(*
SPDX-FileCopyrightText: © 2026 Oleksandr Tiutyk <trofimich@gmail.com>
SPDX-License-Identifier: MIT
License: https://opensource.org/license/mit
*)

(*!
<summary>Creates application-specific activities and conditions for Workflows.CreateElement.</summary>
<description>Invoked in the owning task during configuration. The common creation path registers a successful result.</description>
*)
INTERFACE IWorkflowElementFactory

(*!
<summary>Creates an unregistered element for a recognized qualified PLC type.</summary>
<description>Return zero for an unknown type. For a recognized type return one fresh, unattached dynamic element
associated with workflow. Transfer exclusive ownership on return. On failure clean up before propagating;
a failed allocation must raise terminal OOM. Do not register or publish the element in this callback.</description>
<param name="typeName">Case-sensitive namespace and PLC type name.</param>
<param name="workflow">Prospective owner supplied to the node constructor.</param>
*)
METHOD CreateElement : IWorkflowElement
VAR_INPUT
	typeName : STRING(255);
	workflow : IWorkflow;
END_VAR
END_METHOD

END_INTERFACE

(* stored: Version 1.1.0.1
   Itf IWorkflowElementFactory: Id {9cc421ef-b32d-4108-a997-7db327b6a34b}
   Method CreateElement: Id {ea05d59e-6fe1-4e7d-a1c5-4b27528d95d3} *)
